Fanuc KAREL source: KB00120.KL

PROGRAM KB00120
%NOLOCKGROUP
%ENVIRONMENT MIR
VAR
  P1: POSITION
  P2: POSITION
  P3: INTEGER
  RESULT: XYZWPREXT
BEGIN
  P3 = 1
  RESULT = MIRROR(P1, P2, P3)
END KB00120
